// TIA Portal V15.1 export
// export: Created 2026-11-01T21:38:58.4195394Z, ExportSetting WithDefaults, DisplayName Totally Integrated Automation Portal, DisplayVersion V15.1, DisplayName TIA Portal Openness, DisplayVersion V15.1, DisplayName STEP 7 Professional, DisplayVersion V15.1, DisplayName WinCC Professional, DisplayVersion V15.1
Screen "Root screen"  480x272, Number=1, Template=Template_1
  ScreenLayer 
    TextField "HmiScreenItemData" at 48,122 size 384x22  Text="Welcome to HMI_1 (KTP400 Comfort)!"
